ADAPTER vcm_control (* Adapter Interface *)
  (* Standard: 61499-1 *)
  (* Version 0.0, 10/23/2026, macie, Schneider Electric *)
  PACKAGE Main;
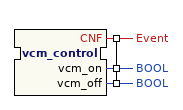
  EVENT_OUTPUT
    CNF WITH vcm_on, vcm_off; (* Confirmation from Plug *)
  END_EVENT
  VAR_OUTPUT
    vcm_on : BOOL; (* Confirmation Data from Plug *)
    vcm_off : BOOL; (* Indication Data from Plug *)
  END_VAR
  SERVICE SOCKET/PLUG
    SEQUENCE request_confirm
      SOCKET.REQ(REQD) -> PLUG.REQ(REQD);
      PLUG.CNF(vcm_on) -> SOCKET.CNF(vcm_on);
    END_SEQUENCE
    SEQUENCE indication_response
      PLUG.IND(vcm_off) -> SOCKET.IND(vcm_off);
      SOCKET.RSP(RSPD) -> PLUG.RSP(RSPD);
    END_SEQUENCE
  END_SERVICE
END_ADAPTER
